FUNCTION_BLOCK FB 7
BEGIN
NETWORK
TITLE = Parsed, but not compiled yet
      A(
      O     I 0.0
      O     I 0.1
      )
      A     DB1.DBX 0.0
      =     Q 0.0
      L     TRUE
END_FUNCTION_BLOCK
